// TIA Portal V21 export
// export: Created 2026-11-08T20:55:21.0056641Z, ExportSetting WithDefaults, DisplayName Totally Integrated Automation Portal, DisplayVersion V21 Update 3, DisplayName STEP 7 Professional, DisplayVersion V21 Update 3, DisplayName STEP 7 Safety, DisplayVersion V21, DisplayName Tech WebApplication, DisplayVersion V21, DisplayName WinCC Basic/Comfort/Advanced, DisplayVersion V21 Update 3, DisplayName WinCC Unified, DisplayVersion V21 Update 3
PlcWatchTable "WT_Test"
  PlcWatchTableEntry ""Tag_Bool_1""  DisplayFormat=Bool, ModifyTrigger=Permanent, MonitorTrigger=Permanent
